FUNCTION_BLOCK F_Gate_Tests EXTENDS TcUnit.FB_TestSuite

Test_ReturnsTrueAndResetsFlag();
Test_ReturnsFalseWhenFlagClear();

METHOD PRIVATE Test_ReturnsTrueAndResetsFlag
VAR
  flag : BOOL;
  result : BOOL;
END_VAR
TcUnit.TEST(__POUNAME());

// arrange
flag := TRUE;

// act
result := F_Gate(flag);

// assert
AssertTrue(Condition := result, Message := 'returns the flag as it was');
AssertFalse(Condition := flag, Message := 'flag reset by the call');

TEST_FINISHED_NAMED(__POUNAME());
END_METHOD

METHOD PRIVATE Test_ReturnsFalseWhenFlagClear
VAR
  flag : BOOL;
  result : BOOL;
END_VAR
TcUnit.TEST(__POUNAME());

// arrange
flag := FALSE;

// act
result := F_Gate(flag);

// assert
AssertFalse(Condition := result, Message := 'clear flag reads FALSE');
AssertFalse(Condition := flag, Message := 'flag stays clear');

TEST_FINISHED_NAMED(__POUNAME());
END_METHOD

END_FUNCTION_BLOCK

(* stored: Version 1.1.0.1, ProductVersion 3.1.4026.22
   POU F_Gate_Tests: Id {070a938d-e118-41b4-8cee-83d1543a7f39}, SpecialFunc None
   Method Test_ReturnsTrueAndResetsFlag: Id {3b4d9a46-659d-4e6d-b210-689ae10b2875}
   Method Test_ReturnsFalseWhenFlagClear: Id {86ba9325-14ee-4e08-bf33-12d87f686ec0} *)
